(* CoDeSys 2.3 export: ld.exp *)

(* POU PLC_LD_PRG_TR, LD *)
PROGRAM PLC_LD_PRG_TR
VAR
END_VAR
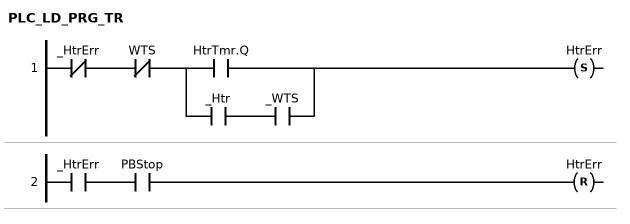
_LD_ (* Ladder Diagram *)
NETWORK 1
	[/_HtrErr] - [/WTS] - { [HtrTmr.Q] | [_Htr] - [_WTS] } --- (S HtrErr)
NETWORK 2
	[_HtrErr] - [PBStop] --- (R HtrErr)
_END_LD_
(* the same logic as Structured Text *)
(* Network 1 *)
IF NOT _HtrErr AND NOT WTS AND (HtrTmr.Q OR _Htr AND _WTS) THEN HtrErr := TRUE; END_IF;
(* Network 2 *)
IF _HtrErr AND PBStop THEN HtrErr := FALSE; END_IF;
END_PROGRAM
